(*
SPDX-FileCopyrightText: © 2026 Oleksandr Tiutyk <trofimich@gmail.com>
SPDX-License-Identifier: MIT
License: https://opensource.org/license/mit
*)

(*!
<summary>
Beckhoff EP2624_0002: 4-channel relay output EtherCAT Box (25 V AC / 30 V DC, make/NO contact, M12).
</summary>
<description>
Process image mapping structure for the EP2624_0002 EtherCAT Box IP67 module with 4 discrete outputs.
The relay ratings are 0.5 A AC at 25 V AC and 2 A DC at 30 V DC; this is not a 230 V AC relay module.
When used for I/O, link located fields or their containing buffers to the matching selected PDOs.
The record is not a packed wire buffer; compiler padding is not part of the device specification.
Unlinked/default values do not prove valid I/O. The caller evaluates bus/channel validity before use.
Use one owner task per instance and externally synchronize other access; multi-field snapshots are not atomic.
Copies store data without creating hardware links. Keep borrowed field references valid while consumers are bound.
This passive record performs no validation, synchronization, configuration or protocol advancement.
</description>
*)
TYPE EP2624_0002 :
STRUCT
	Ch1 AT %Q* : BOOL;
	Ch2 AT %Q* : BOOL;
	Ch3 AT %Q* : BOOL;
	Ch4 AT %Q* : BOOL;
END_STRUCT
END_TYPE

(* stored: Version 1.1.0.1, ProductVersion 3.1.4026.20
   DUT EP2624_0002: Id {80bf3a2b-e4fa-42d9-88b8-237d5ba38585} *)
